Omron CX-Programmer project NewProject (CX-Programmer 9.75)

# PLC NewPLC1: CP1E N30

## Global symbols (name address type ; comment)
0.00 BOOL  ; S1
0.01 BOOL  ; SENSOR
0.02 BOOL  ; S2
0.03 BOOL  ; S3
0.04 BOOL  ; TOR
0.05 BOOL  ; S3
0.06 BOOL  ; TOR
100.00 BOOL  ; H3
100.01 BOOL  ; H1
100.02 BOOL  ; H2
100.03 BOOL  ; PINTU BUKA
100.04 BOOL  ; PINTU TUTUP
100.05 BOOL  ; H4
100.06 BOOL  ; PENGUNCI
10.00 BOOL  ; mulai
T000 BOOL  ; TIMER PINTU KEBUKA
T001 BOOL  ; LAMPU MATI
T002 BOOL  ; LAMPU NYALA

## Program NewProgram1 (cyclic task 0)

### Section Section1

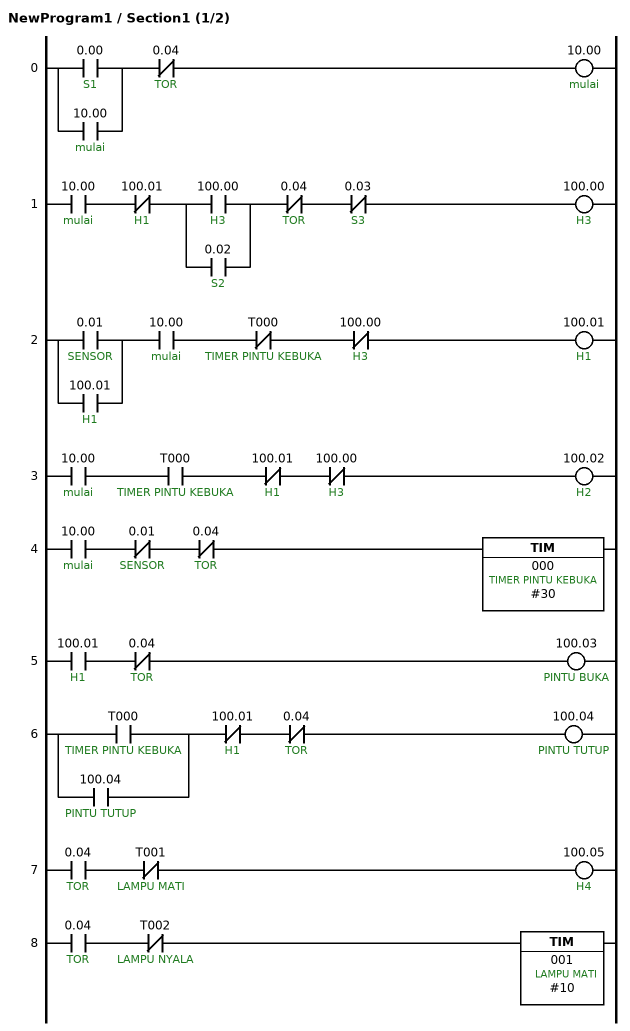
; rung 0
LD 0.00  ; S1
OR 10.00  ; mulai
ANDNOT 0.04  ; TOR
OUT 10.00  ; mulai
; rung 1
LD 10.00  ; mulai
ANDNOT 100.01  ; H1
LD 100.00  ; H3
OR 0.02  ; S2
ANDLD
ANDNOT 0.04  ; TOR
ANDNOT 0.03  ; S3
OUT 100.00  ; H3
; rung 2
LD 0.01  ; SENSOR
OR 100.01  ; H1
AND 10.00  ; mulai
ANDNOT T000  ; TIMER PINTU KEBUKA
ANDNOT 100.00  ; H3
OUT 100.01  ; H1
; rung 3
LD 10.00  ; mulai
AND T000  ; TIMER PINTU KEBUKA
ANDNOT 100.01  ; H1
ANDNOT 100.00  ; H3
OUT 100.02  ; H2
; rung 4
LD 10.00  ; mulai
ANDNOT 0.01  ; SENSOR
ANDNOT 0.04  ; TOR
TIM 000 #30  ; TIMER PINTU KEBUKA
; rung 5
LD 100.01  ; H1
ANDNOT 0.04  ; TOR
OUT 100.03  ; PINTU BUKA
; rung 6
LD T000  ; TIMER PINTU KEBUKA
OR 100.04  ; PINTU TUTUP
ANDNOT 100.01  ; H1
ANDNOT 0.04  ; TOR
OUT 100.04  ; PINTU TUTUP
; rung 7
LD 0.04  ; TOR
ANDNOT T001  ; LAMPU MATI
OUT 100.05  ; H4
; rung 8
LD 0.04  ; TOR
ANDNOT T002  ; LAMPU NYALA
TIM 001 #10  ; LAMPU MATI

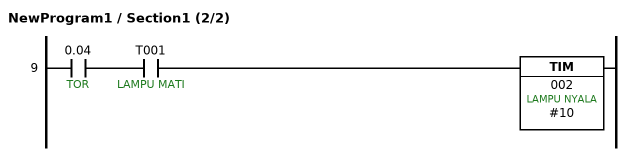
; rung 9
LD 0.04  ; TOR
AND T001  ; LAMPU MATI
TIM 002 #10  ; LAMPU NYALA

### Section END
; rung 0
END(001)